TYPE ST_OperationButtons :
STRUCT
	iActOperation	: E_OperationButtons;
	bSetPause		: BOOL;
	bSetPlay		: BOOL;
	bResetError		: BOOL;
	bStopResetAll	: BOOL;
	bPauseOnDelayed	: BOOL;
	
	bStateSafe_mode : BOOL:=TRUE;
	
	b_rt_Pause		: BOOL;
	b_rt_Play		: BOOL;	

	eModeZone		: E_ModeZone;
	sModeZone		: STRING;
	iPauseHistory	: INT;
	
	iActModeState	: E_WorkingMode; //just for reference stete not for change 
END_STRUCT
END_TYPE

(* stored: Version 1.1.0.1, ProductVersion 3.1.4024.13
   DUT ST_OperationButtons: Id {4f87e27c-78f9-401b-a77e-badff054011e} *)
